(* CODESYS project OperationalMode.xml

Project tree, tasks and I/O mapping:
  visualisation OperationalMode
*)

// /OperationalMode
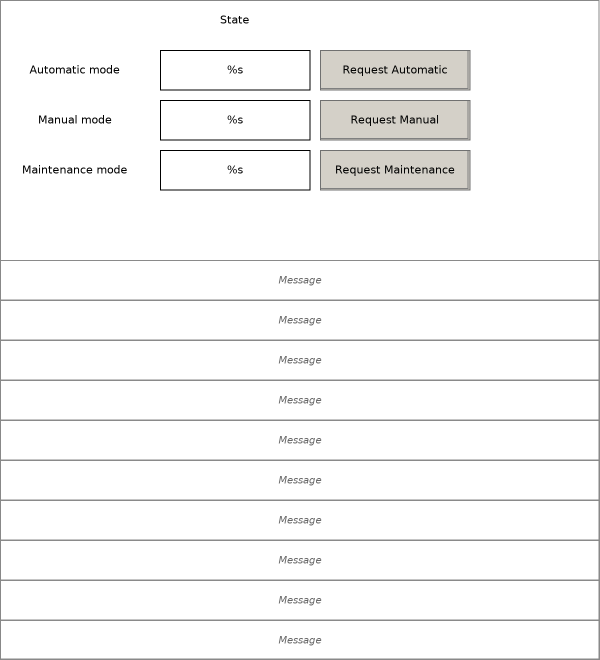
VISUALIZATION OperationalMode  // 600x660
    Button (320,50 150x40), "Request Automatic"
        tap GVL_Project.fbProject._fbModeController._btnRequestAutomatic.xbtn
    Button (320,100 150x40), "Request Manual"
        tap GVL_Project.fbProject._fbModeController._btnRequestManual.xbtn
    Button (320,150 150x40), "Request Maintenance"
        tap GVL_Project.fbProject._fbModeController._btnRequestMaintenance.xbtn
    Rectangle (0,50 150x40), "Automatic mode"
    Rectangle (0,100 150x40), "Manual mode"
    Rectangle (0,150 150x40), "Maintenance mode"
    Rectangle (160,50 150x40), "%s", text variable: GVL_Project.fbProject._fbModeAutomatic._eState
    Rectangle (160,100 150x40), "%s", text variable: GVL_Project.fbProject._fbModeManual._eState
    Rectangle (160,150 150x40), "%s", text variable: GVL_Project.fbProject._fbModeMaintenance._eState
    Rectangle (160,0 150x40), "State"
    Frame (0,260 600x40)
        shows Message(scMessage := GVL_Project.fbProject._fbModeController._ascMessages[1])
    Frame (0,300 600x40)
        shows Message(scMessage := GVL_Project.fbProject._fbModeController._ascMessages[2])
    Frame (0,340 600x40)
        shows Message(scMessage := GVL_Project.fbProject._fbModeController._ascMessages[3])
    Frame (0,380 600x40)
        shows Message(scMessage := GVL_Project.fbProject._fbModeController._ascMessages[4])
    Frame (0,420 600x40)
        shows Message(scMessage := GVL_Project.fbProject._fbModeController._ascMessages[5])
    Frame (0,460 600x40)
        shows Message(scMessage := GVL_Project.fbProject._fbModeController._ascMessages[6])
    Frame (0,500 600x40)
        shows Message(scMessage := GVL_Project.fbProject._fbModeController._ascMessages[7])
    Frame (0,540 600x40)
        shows Message(scMessage := GVL_Project.fbProject._fbModeController._ascMessages[8])
    Frame (0,580 600x40)
        shows Message(scMessage := GVL_Project.fbProject._fbModeController._ascMessages[9])
    Frame (0,620 600x40)
        shows Message(scMessage := GVL_Project.fbProject._fbModeController._ascMessages[10])
END_VISUALIZATION
